// TIA Portal V20 export
// export: Created 2026-10-20T18:54:55.9388741Z, ExportSetting None, DisplayName Totally Integrated Automation Portal, DisplayVersion V20 Update 6, DisplayName TIA Portal Openness, DisplayVersion V20 Update 6, DisplayName TIA Portal Version Control Interface, DisplayVersion V20 Update 6, DisplayName SINAMICS Startdrive Advanced, DisplayVersion V20 SP1, DisplayName SINAMICS Startdrive G130, G150, S120, S150, SINAMICS MV, G220, S200, S210, DisplayVersion V20 SP1, DisplayName SINAMICS Startdrive G110M, G120, G120C, G120D, G120P, G115D, DisplayVersion V20 SP1, DisplayName STEP 7 Professional, DisplayVersion V20 Update 6, DisplayName STEP 7 Safety, DisplayVersion V20 Update 2, DisplayName WinCC Basic/Comfort/Advanced, DisplayVersion V20 Update 6, DisplayName WinCC Unified, DisplayVersion V20 Update 6
VAR_GLOBAL   // PLC tag table "IO_Encoders_2"
   "AE_Control_Word_1(2)" AT %QW210 : UInt;   // 11, 9, 8, 6 … 0 - Reserved / 7 - Fault acknowledge / 10 - Control by PLC / 15...12 - Master’s Sign-of-Life (not relevant)
   "AE_Control_Word_2(2)" AT %QW212 : UInt;   // 10 … 0 - Reserved / 11 - Preset mode / 12 - Activate preset value / 13 - Request for the absolute position value / 14 - Activate park mode / 15 - Acknowledging a sensor error
   "AE_Status_1(2)" AT %IW472 : UInt;   // 8 … 0 - Reserved / 9 - Control requested / 11,10 - Reserved / 15...12 - Encoder’s Sign-of-Life (not relevant)
   "AE_Status_2(2)" AT %IW474 : UInt;   // 9 … 0 - Not supported / 10 - Reserved / 11 - Requirement of error acknowledgement detected / 12 - Status of the Preset function (set/shift of home position executed) / 13 - Transmission of absolute position value / 14 - Park mode activated / 15 - Encoder error
   "AE_Position_1(2)" AT %ID476 : DInt;
   "AE_Position_2(2)" AT %ID480 : DInt;
   "AE_Speed(2)" AT %IW484 : Int;
   "LE_Status(2)" AT %IW271 : UInt;
   "LE_X_Unsafe_Position(2)" AT %ID273 : DInt;
   "LE_Speed(2)" AT %IW277 : Int;   // 0 ...65535
   "LE_Warnings(2)" AT %IW279 : Int;
END_VAR
